(* PLC project g_elevator_door_clean, Anonymous Benchmark Suite 1.0 *)
(* stored: creationDateTime 2026-07-09T00:00:00 *)

PROGRAM g_elevator_door_clean
  VAR_INPUT
    open_req : BOOL;
    move_req : BOOL;
    at_floor : BOOL;
    maint : BOOL;
  END_VAR
  VAR_OUTPUT
    door_open : BOOL;
    drive : BOOL;
  END_VAR

(* LD diagram, written out as Structured Text *)
door_open := NOT move_req AND open_req AND at_floor;
drive := move_req;
END_PROGRAM

CONFIGURATION Config0
  RESOURCE Res0 ON PLC
    TASK tcyclic(INTERVAL := T#10ms, PRIORITY := 0);
    PROGRAM inst0 WITH tcyclic : g_elevator_door_clean;
  END_RESOURCE
END_CONFIGURATION
